Staubli VAL3: do_CASE.pgx

public program do_CASE(string x_sKey, num x_nIndex)
  local num l_nValue
  local string l_sProg
  local string l_sType
begin
  l_nValue=progTemp:pProgItem[x_sKey].pProgTemplate[x_nIndex].sSwitchItem.nSwitchValue
  l_sProg=progTemp:pProgItem[x_sKey].pProgTemplate[x_nIndex].sSwitchItem.sIOValue
  l_sType=progTemp:pProgItem[x_sKey].pProgTemplate[x_nIndex].sTRAJname
  if l_nValue==rs:nSetSwitchValue
    switch l_sType
      case "PROG"
        call makeTraj(l_sProg)
      break
      case "TRAJ"
        call trajectory:makeTraj(l_sProg)
      break
    endSwitch

    rs:nSetSwitchValue=0
    rs:bInSwitch=false
  endIf

end
